(* IEC 61131-3 sources: llm-plc-st-eval/data/definitivo/gemini-3.1-pro-preview/B1/zero_shot, 3 files *)

(* ---- ejec_1.st ---- *)
```iecst
FUNCTION_BLOCK FB_Motor
VAR_INPUT
    btnMarcha : BOOL; // Botón de marcha (TRUE = pulsado)
    btnParo   : BOOL; // Botón de paro (TRUE = pulsado)
    btnEmerg  : BOOL; // Paro de emergencia (TRUE = pulsado)
END_VAR

VAR_OUTPUT
    motorOn   : BOOL; // Estado del motor (TRUE = encendido)
END_VAR

VAR
    rtMarcha  : R_TRIG; // Detector de flanco ascendente
END_VAR

// Detectar flanco ascendente de la marcha para evitar rearranque automático
// si el botón se mantiene pulsado tras un paro de emergencia.
rtMarcha(CLK := btnMarcha);

// Lógica de control (Enclavamiento)
// Prioridad a las señales de paro (btnParo y btnEmerg)
motorOn := (rtMarcha.Q OR motorOn) AND NOT btnParo AND NOT btnEmerg;

END_FUNCTION_BLOCK
```

(* ---- ejec_2.st ---- *)
```iecst
FUNCTION_BLOCK FB_Motor
VAR_INPUT
    btnMarcha : BOOL; // Botón de arranque (TRUE = arrancar)
    btnParo   : BOOL; // Botón de paro normal (TRUE = detener)
    btnEmerg  : BOOL; // Botón de paro de emergencia (TRUE = detener)
END_VAR

VAR_OUTPUT
    motorOn   : BOOL; // Señal de control hacia el contactor del motor
END_VAR

VAR
    flancoMarcha : R_TRIG; // Detector de flanco para el botón de marcha
END_VAR

// Detectar el flanco de subida de la señal de marcha.
// Esto garantiza que el motor no rearranque automáticamente si el
// botón de marcha se mantiene presionado tras un paro de emergencia.
flancoMarcha(CLK := btnMarcha);

// Lógica de control:
// Enclavamiento del motor (flancoMarcha.Q OR motorOn)
// condicionado a que no haya ninguna señal de paro activa.
// El paro y la emergencia tienen prioridad sobre el arranque.
motorOn := (flancoMarcha.Q OR motorOn) AND NOT btnParo AND NOT btnEmerg;

END_FUNCTION_BLOCK
```

(* ---- ejec_3.st ---- *)
```iecst
FUNCTION_BLOCK FB_Motor
VAR_INPUT
    btnMarcha : BOOL; // TRUE al pulsar para arrancar
    btnParo   : BOOL; // TRUE al pulsar para detener
    btnEmerg  : BOOL; // TRUE al activar el paro de emergencia
END_VAR

VAR_OUTPUT
    motorOn   : BOOL; // Estado del motor (TRUE = Encendido)
END_VAR

VAR
    rtMarcha  : R_TRIG; // Detector de flanco de subida para el botón de marcha
END_VAR

// Detección de flanco ascendente para evitar el rearranque automático
// si el botón de marcha se mantiene pulsado tras una emergencia.
rtMarcha(CLK := btnMarcha);

// Lógica de control: Enclavamiento con paro dominante.
// El motor se enciende con el flanco de marcha y se mantiene (motorOn).
// Se detiene inmediatamente si btnParo o btnEmerg son TRUE.
motorOn := (motorOn OR rtMarcha.Q) AND NOT btnParo AND NOT btnEmerg;

END_FUNCTION_BLOCK
```
